Fanuc KAREL source: KA00170.KL

PROGRAM KA00170
%NOLOCKGROUP
VAR
  SRC: ARRAY[4] OF BOOLEAN
  DST: ARRAY[4] OF XYZWPR
BEGIN
  DST = SRC
END KA00170
